(* IEC 61131-3 sources: llm-plc-st-eval/data/processed_v2_primera/claude-sonnet-4-6/B6/few_shot, 3 files *)

(* ---- ejec_1.st ---- *)
FUNCTION_BLOCK FB_Baliza
VAR_INPUT
    alarma : BOOL; (* Condicion de alarma activa *)
END_VAR
VAR_OUTPUT
    lampara : BOOL; (* Lampara de baliza *)
END_VAR
VAR
    tOn  : TON; (* Temporizador fase encendida *)
    tOff : TON; (* Temporizador fase apagada *)
    bParpadeo : BOOL; (* Estado interno del parpadeo *)
END_VAR

(* Sin alarma: lampara apagada y temporizadores reiniciados *)
IF NOT alarma THEN
    bParpadeo := FALSE;
    tOn(IN  := FALSE, PT := T#1S);
    tOff(IN := FALSE, PT := T#1S);
ELSE
    (* Fase encendida: activa tOn mientras bParpadeo es TRUE *)
    tOn(IN := bParpadeo, PT := T#1S);

    (* Fase apagada: activa tOff cuando tOn ha completado *)
    tOff(IN := tOn.Q, PT := T#1S);

    (* Al completar tOff, reiniciar ciclo volviendo a fase encendida *)
    IF tOff.Q THEN
        bParpadeo := FALSE; (* Fuerza reinicio de tOn en el proximo ciclo *)
    END_IF;

    (* Arranque del primer ciclo o reinicio tras fase apagada *)
    IF NOT tOn.IN AND NOT tOff.IN THEN
        bParpadeo := TRUE;
    END_IF;
END_IF;

(* La lampara sigue el estado interno de parpadeo *)
lampara := bParpadeo AND alarma;
END_FUNCTION_BLOCK

(* ---- ejec_2.st ---- *)
FUNCTION_BLOCK FB_Baliza
VAR_INPUT
    alarma : BOOL; (* Condicion de alarma activa *)
END_VAR
VAR_OUTPUT
    lampara : BOOL; (* Lampara de baliza *)
END_VAR
VAR
    tOn  : TON; (* Temporizador fase encendida *)
    tOff : TON; (* Temporizador fase apagada *)
    parpadeo : BOOL; (* Estado interno de parpadeo *)
END_VAR

(* Sin alarma: lampara apagada y temporizadores reiniciados *)
IF NOT alarma THEN
    parpadeo := FALSE;
    tOn(IN  := FALSE, PT := T#1S);
    tOff(IN := FALSE, PT := T#1S);
ELSE
    (* Fase encendida: activa tOn mientras parpadeo=TRUE *)
    tOn(IN := parpadeo, PT := T#1S);

    (* Fase apagada: activa tOff cuando tOn expira *)
    tOff(IN := tOn.Q, PT := T#1S);

    (* Al expirar tOff, reinicia el ciclo volviendo a encender *)
    IF tOff.Q THEN
        parpadeo := FALSE; (* Fuerza reinicio de tOn en el proximo ciclo *)
    END_IF;

    (* Inicia el ciclo si parpadeo esta apagado y tOff no esta corriendo *)
    IF NOT parpadeo AND NOT tOn.Q AND NOT tOff.IN THEN
        parpadeo := TRUE;
    END_IF;
END_IF;

(* La lampara sigue el estado de parpadeo solo durante alarma *)
lampara := alarma AND parpadeo;
END_FUNCTION_BLOCK

(* ---- ejec_3.st ---- *)
FUNCTION_BLOCK FB_Baliza
VAR_INPUT
    alarma : BOOL; (* Condicion de alarma activa *)
END_VAR
VAR_OUTPUT
    lampara : BOOL; (* Lampara de baliza *)
END_VAR
VAR
    tOn  : TON; (* Temporizador fase encendida *)
    tOff : TON; (* Temporizador fase apagada *)
    parpadeo : BOOL; (* Estado interno de parpadeo *)
END_VAR

(* Sin alarma: lampara apagada y temporizadores reiniciados *)
IF NOT alarma THEN
    parpadeo := FALSE;
    tOn(IN  := FALSE, PT := T#1S);
    tOff(IN := FALSE, PT := T#1S);
ELSE
    (* Fase encendida: activa tOn mientras parpadeo = TRUE *)
    tOn(IN := parpadeo, PT := T#1S);

    (* Al completarse tOn, pasa a fase apagada *)
    IF tOn.Q THEN
        parpadeo := FALSE;
        tOn(IN := FALSE, PT := T#1S); (* Reinicia tOn *)
    END_IF;

    (* Fase apagada: activa tOff mientras parpadeo = FALSE *)
    tOff(IN := NOT parpadeo, PT := T#1S);

    (* Al completarse tOff, pasa a fase encendida *)
    IF tOff.Q THEN
        parpadeo := TRUE;
        tOff(IN := FALSE, PT := T#1S); (* Reinicia tOff *)
    END_IF;
END_IF;

(* La lampara sigue el estado de parpadeo solo si hay alarma *)
lampara := alarma AND parpadeo;
END_FUNCTION_BLOCK
